{attribute 'qualified_only'}
{attribute 'strict'}
{attribute 'to_string'}
TYPE E_ModuleMode :
(
	Manual 			:= 0,
	Automatic		:= 1,
	LocalControl 	:= 2, //bypass external control
	DryCycle		:= 3
) INT;
END_TYPE

(* stored: Version 1.1.0.1, ProductVersion 3.1.4024.12
   DUT E_ModuleMode: Id {01603684-8e59-4484-9a93-4730c1d274b4} *)
